(*~
	<docu>
		<summary>
			Writes a little-endian WORD at inOffset.
		</summary>
	</docu>
~*)
FUNCTION TcoAteqG6_SetWord_v_3_5_x : BOOL
VAR_INPUT
	inOffset : INT;
	inValue : WORD;
END_VAR
VAR_IN_OUT
	inoImage : ARRAY[0..255] OF BYTE;
END_VAR

inoImage[inOffset] := WORD_TO_BYTE(inValue AND 16#00FF);
inoImage[inOffset + 1] := WORD_TO_BYTE(SHR(inValue, 8));
TcoAteqG6_SetWord_v_3_5_x := TRUE;

END_FUNCTION

(* stored: Version 1.1.0.1, ProductVersion 3.1.4024.12
   POU TcoAteqG6_SetWord_v_3_5_x: Id {3d788cd7-f3be-43c0-816f-e80fd7b3bfcb}, SpecialFunc None *)
